// TIA Portal V20 export
// export: Created 2026-10-12T05:42:29.8184034Z, ExportSetting WithDefaults, DisplayName Totally Integrated Automation Portal, DisplayVersion V20, DisplayName TIA Portal Openness, DisplayVersion V20, DisplayName TIA Portal Teamcenter Gateway, DisplayVersion V20, DisplayName TIA Portal Version Control Interface, DisplayVersion V20, DisplayName SINAMICS Startdrive Advanced, DisplayVersion V20 SP1 Update 2, DisplayName SINAMICS Startdrive G110M, G120, G120C, G120D, G120P, G115D, DisplayVersion V20 SP1 Update 2, DisplayName SINAMICS Startdrive G130, G150, S120, S150, SINAMICS MV, G220, S200, S210, DisplayVersion V20 SP1 Update 2, DisplayName STEP 7 Professional, DisplayVersion V20, DisplayName STEP 7 Safety, DisplayVersion V20, DisplayName WinCC Basic/Comfort/Advanced, DisplayVersion V20, DisplayName WinCC Professional, DisplayVersion V20, DisplayName WinCC Unified, DisplayVersion V20
FUNCTION "FRK_AccessCrcNumber" : DWord   // FC49, SCL
{ S7_Optimized_Access := 'TRUE' }
VERSION : 0.1
// stored: AutoNumber true, IsIECCheckEnabled false, SetENOAutomatically false, UDAEnableTagReadback false
   VAR_INPUT
      Previous : DWord;
      Value : UDInt;
   END_VAR
   VAR_TEMP
      Index : Int;
      Work : DWord;
   END_VAR
BEGIN

   #Work := #Previous;
   FOR #Index := 0 TO 3 DO
       #Work := "FRK_AccessCrcByte"(Previous := #Work, Value := DWORD_TO_BYTE(SHR(IN := UDINT_TO_DWORD(#Value), N := INT_TO_UINT(#Index * 8))));
   END_FOR;
   #FRK_AccessCrcNumber := #Work;
END_FUNCTION
